KUKA KRL program: MAIN_1.src, MAIN_1.dat

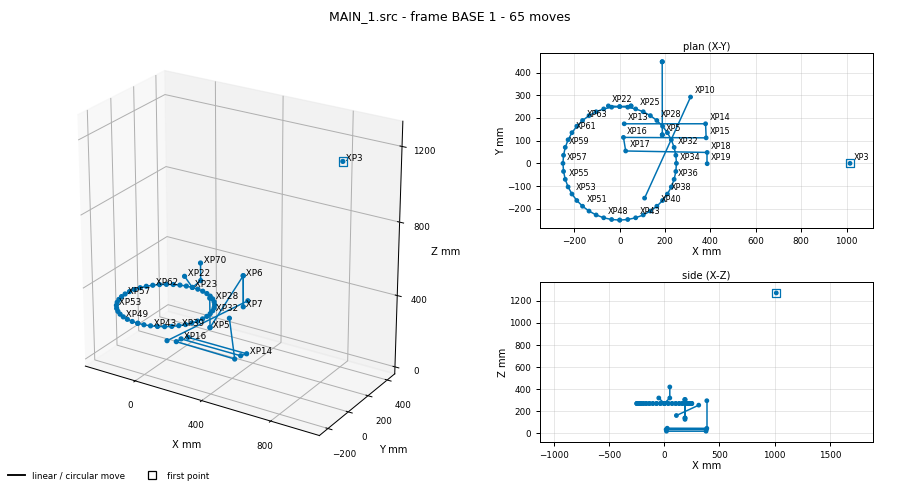
[picture p0: tool path of MAIN_1.src in frame BASE 1, 65 of 76 moves have a stored position in this frame; points joined in program order, loops and branches not executed]
--- MAIN_1.src ---
&ACCESS RVP
&REL 1
&COMMENT Generated by RoboDK
&PARAM TEMPLATE = C:\KRC\Roboter\Template\vorgabe
&PARAM EDITMASK = *
DEF MAIN_1 ( )
;FOLD INI
BAS (#INITMOV,0 )
;ENDFOLD (INI)

;FOLD STARTPOS
$BWDSTART = FALSE
PDAT_ACT = {VEL 50,ACC 100,APO_DIST 10}
BAS(#PTP_DAT)
FDAT_ACT = {TOOL_NO 0,BASE_NO 0,IPO_FRAME #BASE}
BAS (#FRAMES)
BAS (#VEL_PTP,50)
;ENDFOLD


;FOLD SET DEFAULT SPEED
$VEL.CP=0.2
BAS(#VEL_PTP,50)
BAS(#TOOL,0)
BAS(#BASE,0)
;ENDFOLD

;FOLD PTP FIRST POSITION
$BWDSTART = FALSE
PDAT_ACT = {VEL 50,ACC 100,APO_DIST 10}
FDAT_ACT = {TOOL_NO 0,BASE_NO 0,IPO_FRAME #BASE}
BAS(#FRAMES)
$ADVANCE = 5
;ENDFOLD

PTP $AXIS_ACT ; skip BCO quickly

; Program generated by RoboDK v5.6.9 for RoboDK Industrial on 26/02/2024 09:58:20
; Using nominal kinematics.
;FOLD PTP P1 Vel=100.000 % PDAT1 Tool[1] Base[1];%{PE}%R 8.3.42,%MKUKATPBASIS,%CMOVE,%VPTP,%P 1:PTP, 2:P1, 3:, 5:100, 7:PDAT1
$BWDSTART=FALSE
PDAT_ACT=PPDAT1
FDAT_ACT=FP1
BAS(#PTP_PARAMS,100)
PTP XP1 C_PTP
;ENDFOLD
;FOLD PTP P2 Vel=100.000 % PDAT2 Tool[1] Base[1];%{PE}%R 8.3.42,%MKUKATPBASIS,%CMOVE,%VPTP,%P 1:PTP, 2:P2, 3:, 5:100, 7:PDAT2
$BWDSTART=FALSE
PDAT_ACT=PPDAT2
FDAT_ACT=FP2
BAS(#PTP_PARAMS,100)
PTP XP2 C_PTP
;ENDFOLD
;FOLD LIN P3 Vel=1.000 m/s CPDAT3 Tool[1] Base[1];%{PE}%R 8.3.42,%MKUKATPBASIS,%CMOVE,%VLIN,%P 1:LIN, 2:P3, 3:, 5:1, 7:CPDAT3
$BWDSTART=FALSE
LDAT_ACT=LCPDAT3
FDAT_ACT=FP3
BAS(#CP_PARAMS,1.000)
LIN XP3 C_DIS
;ENDFOLD
$OUT[5]=TRUE
$OUT[5]=TRUE
$OUT[5]=0.5
$OUT[5]=true
$ANOUT[5]=TRUE
$ANOUT[5]=TRUE
$ANOUT[5]=0.5
$ANOUT[5]=true
var=val
var=val
WAIT FOR ($IN[5]==TRUE)
WAIT FOR ($IN[5]==TRUE)
WAIT FOR ($IN[5]==0.5)
WAIT FOR ($IN[5]==true)
START_TIMER:
$TIMER_STOP[1]=TRUE
$TIMER_FLAG[1]=FALSE
$TIMER[1]=0.100
$TIMER_STOP[1]=FALSE
WAIT FOR ($IN[5]==TRUE OR $TIMER_FLAG[1])
$TIMER_STOP[1]=TRUE
IF $TIMER_FLAG[1]== TRUE THEN
    HALT ; Timed out!
    GOTO START_TIMER
ENDIF
WAIT FOR (var==val)
START_TIMER:
$TIMER_STOP[1]=TRUE
$TIMER_FLAG[1]=FALSE
$TIMER[1]=0.100
$TIMER_STOP[1]=FALSE
WAIT FOR (var==val OR $TIMER_FLAG[1])
$TIMER_STOP[1]=TRUE
IF $TIMER_FLAG[1]== TRUE THEN
    HALT ; Timed out!
    GOTO START_TIMER
ENDIF
Wait for StrClear($LOOP_MSG[])
$LOOP_CONT = TRUE
$LOOP_MSG[] = "Message"
REMOTE_PROG_CALL_171()
CODE_INSERT_172
; Insert Comment
; ---- Setting reference (Base) ----
$BASE = {FRAME: X 719.013,Y -664.003,Z 0.000,A 0.000,B 0.000,C 0.000}
; --------------------------
; ---- Setting tool (TCP) ----
; TOOL_DATA[1] = {FRAME: X 129.073,Y 0.000,Z 85.477,A 0.000,B 22.849,C 0.000}
$TOOL = {FRAME: X 129.073,Y 0.000,Z 85.477,A 0.000,B 22.849,C 0.000}
; $TOOL = TOOL_DATA[1]
; --------------------------
$ACC.ORI1 = 800.00000
$ACC.ORI2 = 800.00000
$VEL.ORI1 = 500.00000
$VEL.ORI2 = 500.00000
$APO.CPTP = 10
$APO.CDIS = 10.000
;FOLD PTP P4 CONT Vel=100.000 % PDAT4 Tool[1] Base[1];%{PE}%R 8.3.42,%MKUKATPBASIS,%CMOVE,%VPTP,%P 1:PTP, 2:P4, 3:C_PTP, 5:100, 7:PDAT4
$BWDSTART=FALSE
PDAT_ACT=PPDAT4
FDAT_ACT=FP4
BAS(#PTP_PARAMS,100)
PTP XP4 C_PTP
;ENDFOLD
$ACC.CP = 0.20000
$VEL.CP = 0.10000
;FOLD LIN P5 Vel=0.100 m/s CPDAT5 Tool[1] Base[1];%{PE}%R 8.3.42,%MKUKATPBASIS,%CMOVE,%VLIN,%P 1:LIN, 2:P5, 3:, 5:0, 7:CPDAT5
$BWDSTART=FALSE
LDAT_ACT=LCPDAT5
FDAT_ACT=FP5
BAS(#CP_PARAMS,0.100)
LIN XP5 C_DIS
;ENDFOLD
$OUT[5]=TRUE
PICK_PART_111()
$APO.CPTP = 10
$APO.CDIS = 10.000
$ACC.CP = 0.60000
$VEL.CP = 0.30000
; Linear movement using joint targets is not supported. Change the target type to cartesian or use a joint movement.
;FOLD LIN P6 CONT Vel=0.300 m/s CPDAT6 Tool[1] Base[1];%{PE}%R 8.3.42,%MKUKATPBASIS,%CMOVE,%VLIN,%P 1:LIN, 2:P6, 3:C_DIS, 5:0, 7:CPDAT6
$BWDSTART=FALSE
LDAT_ACT=LCPDAT6
FDAT_ACT=FP6
BAS(#CP_PARAMS,0.300)
LIN XP6 C_DIS
;ENDFOLD
$ACC.CP = 0.20000
$VEL.CP = 0.10000
; MoveSearch command not implemented
;FOLD LIN P7 Vel=0.100 m/s CPDAT7 Tool[1] Base[1];%{PE}%R 8.3.42,%MKUKATPBASIS,%CMOVE,%VLIN,%P 1:LIN, 2:P7, 3:, 5:0, 7:CPDAT7
$BWDSTART=FALSE
LDAT_ACT=LCPDAT7
FDAT_ACT=FP7
BAS(#CP_PARAMS,0.100)
LIN XP7 C_DIS
;ENDFOLD
$OUT[5]=FALSE
PLACE_PART_112()
$APO.CPTP = 10
$APO.CDIS = 10.000
;FOLD LIN P8 CONT Vel=0.100 m/s CPDAT8 Tool[1] Base[1];%{PE}%R 8.3.42,%MKUKATPBASIS,%CMOVE,%VLIN,%P 1:LIN, 2:P8, 3:C_DIS, 5:0, 7:CPDAT8
$BWDSTART=FALSE
LDAT_ACT=LCPDAT8
FDAT_ACT=FP8
BAS(#CP_PARAMS,0.100)
LIN XP8 C_DIS
;ENDFOLD
; ---- Setting reference (Base) ----
$BASE = {FRAME: X 577.670,Y 392.250,Z 0.000,A 38.960,B 0.000,C 0.000}
; --------------------------
$APO.CPTP = 25
$APO.CDIS = 25.000
$ACC.ORI1 = 800.00000
$ACC.ORI2 = 800.00000
$VEL.ORI1 = 500.00000
$VEL.ORI2 = 500.00000
$ACC.CP = 0.20000
$VEL.CP = 0.10000
;FOLD PTP P9 CONT Vel=100.000 % PDAT9 Tool[1] Base[1];%{PE}%R 8.3.42,%MKUKATPBASIS,%CMOVE,%VPTP,%P 1:PTP, 2:P9, 3:C_PTP, 5:100, 7:PDAT9
$BWDSTART=FALSE
PDAT_ACT=PPDAT9
FDAT_ACT=FP9
BAS(#PTP_PARAMS,100)
PTP XP9 C_PTP
;ENDFOLD
CIRC {X 430.047,Y 43.774,Z 231.503,A -134.549,B 11.181,C 178.913},{X 109.688,Y -153.222,Z 161.073,A -134.549,B 11.181,C 178.913} C_DIS
; Circular movement using joint targets is not supported. Change the target type to cartesian or use a joint movement.
$ACC.CP = 0.20000
$VEL.CP = 0.10000
;FOLD LIN P10 Vel=0.100 m/s CPDAT10 Tool[1] Base[1];%{PE}%R 8.3.42,%MKUKATPBASIS,%CMOVE,%VLIN,%P 1:LIN, 2:P10, 3:, 5:0, 7:CPDAT10
$BWDSTART=FALSE
LDAT_ACT=LCPDAT10
FDAT_ACT=FP10
BAS(#CP_PARAMS,0.100)
LIN XP10 C_DIS
;ENDFOLD
;FOLD PTP P11 Vel=100.000 % PDAT11 Tool[1] Base[1];%{PE}%R 8.3.42,%MKUKATPBASIS,%CMOVE,%VPTP,%P 1:PTP, 2:P11, 3:, 5:100, 7:PDAT11
$BWDSTART=FALSE
PDAT_ACT=PPDAT11
FDAT_ACT=FP11
BAS(#PTP_PARAMS,100)
PTP XP11 C_PTP
;ENDFOLD
; ---- Setting reference (Base) ----
$BASE = {FRAME: X 0.000,Y 782.714,Z 377.610,A 0.000,B 0.000,C 0.000}
; --------------------------
;FOLD PTP P12 Vel=100.000 % PDAT12 Tool[1] Base[1];%{PE}%R 8.3.42,%MKUKATPBASIS,%CMOVE,%VPTP,%P 1:PTP, 2:P12, 3:, 5:100, 7:PDAT12
$BWDSTART=FALSE
PDAT_ACT=PPDAT12
FDAT_ACT=FP12
BAS(#PTP_PARAMS,100)
PTP XP12 C_PTP
;ENDFOLD
;FOLD LIN P13 Vel=0.100 m/s CPDAT13 Tool[1] Base[1];%{PE}%R 8.3.42,%MKUKATPBASIS,%CMOVE,%VLIN,%P 1:LIN, 2:P13, 3:, 5:0, 7:CPDAT13
$BWDSTART=FALSE
LDAT_ACT=LCPDAT13
FDAT_ACT=FP13
BAS(#CP_PARAMS,0.100)
LIN XP13 C_DIS
;ENDFOLD
;FOLD LIN P14 Vel=0.100 m/s CPDAT14 Tool[1] Base[1];%{PE}%R 8.3.42,%MKUKATPBASIS,%CMOVE,%VLIN,%P 1:LIN, 2:P14, 3:, 5:0, 7:CPDAT14
$BWDSTART=FALSE
LDAT_ACT=LCPDAT14
FDAT_ACT=FP14
BAS(#CP_PARAMS,0.100)
LIN XP14 C_DIS
;ENDFOLD
;FOLD LIN P15 Vel=0.100 m/s CPDAT15 Tool[1] Base[1];%{PE}%R 8.3.42,%MKUKATPBASIS,%CMOVE,%VLIN,%P 1:LIN, 2:P15, 3:, 5:0, 7:CPDAT15
$BWDSTART=FALSE
LDAT_ACT=LCPDAT15
FDAT_ACT=FP15
BAS(#CP_PARAMS,0.100)
LIN XP15 C_DIS
;ENDFOLD
;FOLD LIN P16 Vel=0.100 m/s CPDAT16 Tool[1] Base[1];%{PE}%R 8.3.42,%MKUKATPBASIS,%CMOVE,%VLIN,%P 1:LIN, 2:P16, 3:, 5:0, 7:CPDAT16
$BWDSTART=FALSE
LDAT_ACT=LCPDAT16
FDAT_ACT=FP16
BAS(#CP_PARAMS,0.100)
LIN XP16 C_DIS
;ENDFOLD
;FOLD LIN P17 Vel=0.100 m/s CPDAT17 Tool[1] Base[1];%{PE}%R 8.3.42,%MKUKATPBASIS,%CMOVE,%VLIN,%P 1:LIN, 2:P17, 3:, 5:0, 7:CPDAT17
$BWDSTART=FALSE
LDAT_ACT=LCPDAT17
FDAT_ACT=FP17
BAS(#CP_PARAMS,0.100)
LIN XP17 C_DIS
;ENDFOLD
;FOLD LIN P18 Vel=0.100 m/s CPDAT18 Tool[1] Base[1];%{PE}%R 8.3.42,%MKUKATPBASIS,%CMOVE,%VLIN,%P 1:LIN, 2:P18, 3:, 5:0, 7:CPDAT18
$BWDSTART=FALSE
LDAT_ACT=LCPDAT18
FDAT_ACT=FP18
BAS(#CP_PARAMS,0.100)
LIN XP18 C_DIS
;ENDFOLD
;FOLD LIN P19 Vel=0.100 m/s CPDAT19 Tool[1] Base[1];%{PE}%R 8.3.42,%MKUKATPBASIS,%CMOVE,%VLIN,%P 1:LIN, 2:P19, 3:, 5:0, 7:CPDAT19
$BWDSTART=FALSE
LDAT_ACT=LCPDAT19
FDAT_ACT=FP19
BAS(#CP_PARAMS,0.100)
LIN XP19 C_DIS
;ENDFOLD
;FOLD PTP P20 Vel=100.000 % PDAT20 Tool[1] Base[1];%{PE}%R 8.3.42,%MKUKATPBASIS,%CMOVE,%VPTP,%P 1:PTP, 2:P20, 3:, 5:100, 7:PDAT20
$BWDSTART=FALSE
PDAT_ACT=PPDAT20
FDAT_ACT=FP20
BAS(#PTP_PARAMS,100)
PTP XP20 C_PTP
;ENDFOLD
EVENT_PROG_START_101()
$APO.CPTP = 1
$APO.CDIS = 1.000
$VEL.CP = 1.00000
; ---- Setting reference (Base) ----
$BASE = {FRAME: X 13.637,Y -840.080,Z 0.000,A -90.000,B 0.000,C 0.000}
; --------------------------
; Show Tool 1
;FOLD PTP P21 CONT Vel=100.000 % PDAT21 Tool[1] Base[1];%{PE}%R 8.3.42,%MKUKATPBASIS,%CMOVE,%VPTP,%P 1:PTP, 2:P21, 3:C_PTP, 5:100, 7:PDAT21
$BWDSTART=FALSE
PDAT_ACT=PPDAT21
FDAT_ACT=FP21
BAS(#PTP_PARAMS,100)
PTP XP21 C_PTP
;ENDFOLD
EVENT_PATH_APPROACH_102()
;FOLD LIN P22 CONT Vel=1.000 m/s CPDAT22 Tool[1] Base[1];%{PE}%R 8.3.42,%MKUKATPBASIS,%CMOVE,%VLIN,%P 1:LIN, 2:P22, 3:C_DIS, 5:1, 7:CPDAT22
$BWDSTART=FALSE
LDAT_ACT=LCPDAT22
FDAT_ACT=FP22
BAS(#CP_PARAMS,1.000)
LIN XP22 C_DIS
;ENDFOLD
;FOLD LIN P23 CONT Vel=1.000 m/s CPDAT23 Tool[1] Base[1];%{PE}%R 8.3.42,%MKUKATPBASIS,%CMOVE,%VLIN,%P 1:LIN, 2:P23, 3:C_DIS, 5:1, 7:CPDAT23
$BWDSTART=FALSE
LDAT_ACT=LCPDAT23
FDAT_ACT=FP23
BAS(#CP_PARAMS,1.000)
LIN XP23 C_DIS
;ENDFOLD
EVENT_PATH_START_103()
$VEL.CP = 0.05000
;FOLD LIN P24 CONT Vel=0.050 m/s CPDAT24 Tool[1] Base[1];%{PE}%R 8.3.42,%MKUKATPBASIS,%CMOVE,%VLIN,%P 1:LIN, 2:P24, 3:C_DIS, 5:0, 7:CPDAT24
$BWDSTART=FALSE
LDAT_ACT=LCPDAT24
FDAT_ACT=FP24
BAS(#CP_PARAMS,0.050)
LIN XP24 C_DIS
;ENDFOLD
;FOLD LIN P25 CONT Vel=0.050 m/s CPDAT25 Tool[1] Base[1];%{PE}%R 8.3.42,%MKUKATPBASIS,%CMOVE,%VLIN,%P 1:LIN, 2:P25, 3:C_DIS, 5:0, 7:CPDAT25
$BWDSTART=FALSE
LDAT_ACT=LCPDAT25
FDAT_ACT=FP25
BAS(#CP_PARAMS,0.050)
LIN XP25 C_DIS
;ENDFOLD
;FOLD LIN P26 CONT Vel=0.050 m/s CPDAT26 Tool[1] Base[1];%{PE}%R 8.3.42,%MKUKATPBASIS,%CMOVE,%VLIN,%P 1:LIN, 2:P26, 3:C_DIS, 5:0, 7:CPDAT26
$BWDSTART=FALSE
LDAT_ACT=LCPDAT26
FDAT_ACT=FP26
BAS(#CP_PARAMS,0.050)
LIN XP26 C_DIS
;ENDFOLD
;FOLD LIN P27 CONT Vel=0.050 m/s CPDAT27 Tool[1] Base[1];%{PE}%R 8.3.42,%MKUKATPBASIS,%CMOVE,%VLIN,%P 1:LIN, 2:P27, 3:C_DIS, 5:0, 7:CPDAT27
$BWDSTART=FALSE
LDAT_ACT=LCPDAT27
FDAT_ACT=FP27
BAS(#CP_PARAMS,0.050)
LIN XP27 C_DIS
;ENDFOLD
;FOLD LIN P28 CONT Vel=0.050 m/s CPDAT28 Tool[1] Base[1];%{PE}%R 8.3.42,%MKUKATPBASIS,%CMOVE,%VLIN,%P 1:LIN, 2:P28, 3:C_DIS, 5:0, 7:CPDAT28
$BWDSTART=FALSE
LDAT_ACT=LCPDAT28
FDAT_ACT=FP28
BAS(#CP_PARAMS,0.050)
LIN XP28 C_DIS
;ENDFOLD
;FOLD LIN P29 CONT Vel=0.050 m/s CPDAT29 Tool[1] Base[1];%{PE}%R 8.3.42,%MKUKATPBASIS,%CMOVE,%VLIN,%P 1:LIN, 2:P29, 3:C_DIS, 5:0, 7:CPDAT29
$BWDSTART=FALSE
LDAT_ACT=LCPDAT29
FDAT_ACT=FP29
BAS(#CP_PARAMS,0.050)
LIN XP29 C_DIS
;ENDFOLD
;FOLD LIN P30 CONT Vel=0.050 m/s CPDAT30 Tool[1] Base[1];%{PE}%R 8.3.42,%MKUKATPBASIS,%CMOVE,%VLIN,%P 1:LIN, 2:P30, 3:C_DIS, 5:0, 7:CPDAT30
$BWDSTART=FALSE
LDAT_ACT=LCPDAT30
FDAT_ACT=FP30
BAS(#CP_PARAMS,0.050)
LIN XP30 C_DIS
;ENDFOLD
;FOLD LIN P31 CONT Vel=0.050 m/s CPDAT31 Tool[1] Base[1];%{PE}%R 8.3.42,%MKUKATPBASIS,%CMOVE,%VLIN,%P 1:LIN, 2:P31, 3:C_DIS, 5:0, 7:CPDAT31
$BWDSTART=FALSE
LDAT_ACT=LCPDAT31
FDAT_ACT=FP31
BAS(#CP_PARAMS,0.050)
LIN XP31 C_DIS
;ENDFOLD
;FOLD LIN P32 CONT Vel=0.050 m/s CPDAT32 Tool[1] Base[1];%{PE}%R 8.3.42,%MKUKATPBASIS,%CMOVE,%VLIN,%P 1:LIN, 2:P32, 3:C_DIS, 5:0, 7:CPDAT32
$BWDSTART=FALSE
LDAT_ACT=LCPDAT32
FDAT_ACT=FP32
BAS(#CP_PARAMS,0.050)
LIN XP32 C_DIS
;ENDFOLD
;FOLD LIN P33 CONT Vel=0.050 m/s CPDAT33 Tool[1] Base[1];%{PE}%R 8.3.42,%MKUKATPBASIS,%CMOVE,%VLIN,%P 1:LIN, 2:P33, 3:C_DIS, 5:0, 7:CPDAT33
$BWDSTART=FALSE
LDAT_ACT=LCPDAT33
FDAT_ACT=FP33
BAS(#CP_PARAMS,0.050)
LIN XP33 C_DIS
;ENDFOLD
;FOLD LIN P34 CONT Vel=0.050 m/s CPDAT34 Tool[1] Base[1];%{PE}%R 8.3.42,%MKUKATPBASIS,%CMOVE,%VLIN,%P 1:LIN, 2:P34, 3:C_DIS, 5:0, 7:CPDAT34
$BWDSTART=FALSE
LDAT_ACT=LCPDAT34
FDAT_ACT=FP34
BAS(#CP_PARAMS,0.050)
LIN XP34 C_DIS
;ENDFOLD
;FOLD LIN P35 CONT Vel=0.050 m/s CPDAT35 Tool[1] Base[1];%{PE}%R 8.3.42,%MKUKATPBASIS,%CMOVE,%VLIN,%P 1:LIN, 2:P35, 3:C_DIS, 5:0, 7:CPDAT35
$BWDSTART=FALSE
LDAT_ACT=LCPDAT35
FDAT_ACT=FP35
BAS(#CP_PARAMS,0.050)
LIN XP35 C_DIS
;ENDFOLD
;FOLD LIN P36 CONT Vel=0.050 m/s CPDAT36 Tool[1] Base[1];%{PE}%R 8.3.42,%MKUKATPBASIS,%CMOVE,%VLIN,%P 1:LIN, 2:P36, 3:C_DIS, 5:0, 7:CPDAT36
$BWDSTART=FALSE
LDAT_ACT=LCPDAT36
FDAT_ACT=FP36
BAS(#CP_PARAMS,0.050)
LIN XP36 C_DIS
;ENDFOLD
;FOLD LIN P37 CONT Vel=0.050 m/s CPDAT37 Tool[1] Base[1];%{PE}%R 8.3.42,%MKUKATPBASIS,%CMOVE,%VLIN,%P 1:LIN, 2:P37, 3:C_DIS, 5:0, 7:CPDAT37
$BWDSTART=FALSE
LDAT_ACT=LCPDAT37
FDAT_ACT=FP37
BAS(#CP_PARAMS,0.050)
LIN XP37 C_DIS
;ENDFOLD
;FOLD LIN P38 CONT Vel=0.050 m/s CPDAT38 Tool[1] Base[1];%{PE}%R 8.3.42,%MKUKATPBASIS,%CMOVE,%VLIN,%P 1:LIN, 2:P38, 3:C_DIS, 5:0, 7:CPDAT38
$BWDSTART=FALSE
LDAT_ACT=LCPDAT38
FDAT_ACT=FP38
BAS(#CP_PARAMS,0.050)
LIN XP38 C_DIS
;ENDFOLD
;FOLD LIN P39 CONT Vel=0.050 m/s CPDAT39 Tool[1] Base[1];%{PE}%R 8.3.42,%MKUKATPBASIS,%CMOVE,%VLIN,%P 1:LIN, 2:P39, 3:C_DIS, 5:0, 7:CPDAT39
$BWDSTART=FALSE
LDAT_ACT=LCPDAT39
FDAT_ACT=FP39
BAS(#CP_PARAMS,0.050)
LIN XP39 C_DIS
;ENDFOLD
;FOLD LIN P40 CONT Vel=0.050 m/s CPDAT40 Tool[1] Base[1];%{PE}%R 8.3.42,%MKUKATPBASIS,%CMOVE,%VLIN,%P 1:LIN, 2:P40, 3:C_DIS, 5:0, 7:CPDAT40
$BWDSTART=FALSE
LDAT_ACT=LCPDAT40
FDAT_ACT=FP40
BAS(#CP_PARAMS,0.050)
LIN XP40 C_DIS
;ENDFOLD
;FOLD LIN P41 CONT Vel=0.050 m/s CPDAT41 Tool[1] Base[1];%{PE}%R 8.3.42,%MKUKATPBASIS,%CMOVE,%VLIN,%P 1:LIN, 2:P41, 3:C_DIS, 5:0, 7:CPDAT41
$BWDSTART=FALSE
LDAT_ACT=LCPDAT41
FDAT_ACT=FP41
BAS(#CP_PARAMS,0.050)
LIN XP41 C_DIS
;ENDFOLD
;FOLD LIN P42 CONT Vel=0.050 m/s CPDAT42 Tool[1] Base[1];%{PE}%R 8.3.42,%MKUKATPBASIS,%CMOVE,%VLIN,%P 1:LIN, 2:P42, 3:C_DIS, 5:0, 7:CPDAT42
$BWDSTART=FALSE
LDAT_ACT=LCPDAT42
FDAT_ACT=FP42
BAS(#CP_PARAMS,0.050)
LIN XP42 C_DIS
;ENDFOLD
;FOLD LIN P43 CONT Vel=0.050 m/s CPDAT43 Tool[1] Base[1];%{PE}%R 8.3.42,%MKUKATPBASIS,%CMOVE,%VLIN,%P 1:LIN, 2:P43, 3:C_DIS, 5:0, 7:CPDAT43
$BWDSTART=FALSE
LDAT_ACT=LCPDAT43
FDAT_ACT=FP43
BAS(#CP_PARAMS,0.050)
LIN XP43 C_DIS
;ENDFOLD
;FOLD LIN P44 CONT Vel=0.050 m/s CPDAT44 Tool[1] Base[1];%{PE}%R 8.3.42,%MKUKATPBASIS,%CMOVE,%VLIN,%P 1:LIN, 2:P44, 3:C_DIS, 5:0, 7:CPDAT44
$BWDSTART=FALSE
LDAT_ACT=LCPDAT44
FDAT_ACT=FP44
BAS(#CP_PARAMS,0.050)
LIN XP44 C_DIS
;ENDFOLD
;FOLD LIN P45 CONT Vel=0.050 m/s CPDAT45 Tool[1] Base[1];%{PE}%R 8.3.42,%MKUKATPBASIS,%CMOVE,%VLIN,%P 1:LIN, 2:P45, 3:C_DIS, 5:0, 7:CPDAT45
$BWDSTART=FALSE
LDAT_ACT=LCPDAT45
FDAT_ACT=FP45
BAS(#CP_PARAMS,0.050)
LIN XP45 C_DIS
;ENDFOLD
;FOLD LIN P46 CONT Vel=0.050 m/s CPDAT46 Tool[1] Base[1];%{PE}%R 8.3.42,%MKUKATPBASIS,%CMOVE,%VLIN,%P 1:LIN, 2:P46, 3:C_DIS, 5:0, 7:CPDAT46
$BWDSTART=FALSE
LDAT_ACT=LCPDAT46
FDAT_ACT=FP46
BAS(#CP_PARAMS,0.050)
LIN XP46 C_DIS
;ENDFOLD
;FOLD LIN P47 CONT Vel=0.050 m/s CPDAT47 Tool[1] Base[1];%{PE}%R 8.3.42,%MKUKATPBASIS,%CMOVE,%VLIN,%P 1:LIN, 2:P47, 3:C_DIS, 5:0, 7:CPDAT47
$BWDSTART=FALSE
LDAT_ACT=LCPDAT47
FDAT_ACT=FP47
BAS(#CP_PARAMS,0.050)
LIN XP47 C_DIS
;ENDFOLD
;FOLD LIN P48 CONT Vel=0.050 m/s CPDAT48 Tool[1] Base[1];%{PE}%R 8.3.42,%MKUKATPBASIS,%CMOVE,%VLIN,%P 1:LIN, 2:P48, 3:C_DIS, 5:0, 7:CPDAT48
$BWDSTART=FALSE
LDAT_ACT=LCPDAT48
FDAT_ACT=FP48
BAS(#CP_PARAMS,0.050)
LIN XP48 C_DIS
;ENDFOLD
;FOLD LIN P49 CONT Vel=0.050 m/s CPDAT49 Tool[1] Base[1];%{PE}%R 8.3.42,%MKUKATPBASIS,%CMOVE,%VLIN,%P 1:LIN, 2:P49, 3:C_DIS, 5:0, 7:CPDAT49
$BWDSTART=FALSE
LDAT_ACT=LCPDAT49
FDAT_ACT=FP49
BAS(#CP_PARAMS,0.050)
LIN XP49 C_DIS
;ENDFOLD
;FOLD LIN P50 CONT Vel=0.050 m/s CPDAT50 Tool[1] Base[1];%{PE}%R 8.3.42,%MKUKATPBASIS,%CMOVE,%VLIN,%P 1:LIN, 2:P50, 3:C_DIS, 5:0, 7:CPDAT50
$BWDSTART=FALSE
LDAT_ACT=LCPDAT50
FDAT_ACT=FP50
BAS(#CP_PARAMS,0.050)
LIN XP50 C_DIS
;ENDFOLD
;FOLD LIN P51 CONT Vel=0.050 m/s CPDAT51 Tool[1] Base[1];%{PE}%R 8.3.42,%MKUKATPBASIS,%CMOVE,%VLIN,%P 1:LIN, 2:P51, 3:C_DIS, 5:0, 7:CPDAT51
$BWDSTART=FALSE
LDAT_ACT=LCPDAT51
FDAT_ACT=FP51
BAS(#CP_PARAMS,0.050)
LIN XP51 C_DIS
;ENDFOLD
;FOLD LIN P52 CONT Vel=0.050 m/s CPDAT52 Tool[1] Base[1];%{PE}%R 8.3.42,%MKUKATPBASIS,%CMOVE,%VLIN,%P 1:LIN, 2:P52, 3:C_DIS, 5:0, 7:CPDAT52
$BWDSTART=FALSE
LDAT_ACT=LCPDAT52
FDAT_ACT=FP52
BAS(#CP_PARAMS,0.050)
LIN XP52 C_DIS
;ENDFOLD
;FOLD LIN P53 CONT Vel=0.050 m/s CPDAT53 Tool[1] Base[1];%{PE}%R 8.3.42,%MKUKATPBASIS,%CMOVE,%VLIN,%P 1:LIN, 2:P53, 3:C_DIS, 5:0, 7:CPDAT53
$BWDSTART=FALSE
LDAT_ACT=LCPDAT53
FDAT_ACT=FP53
BAS(#CP_PARAMS,0.050)
LIN XP53 C_DIS
;ENDFOLD
;FOLD LIN P54 CONT Vel=0.050 m/s CPDAT54 Tool[1] Base[1];%{PE}%R 8.3.42,%MKUKATPBASIS,%CMOVE,%VLIN,%P 1:LIN, 2:P54, 3:C_DIS, 5:0, 7:CPDAT54
$BWDSTART=FALSE
LDAT_ACT=LCPDAT54
FDAT_ACT=FP54
BAS(#CP_PARAMS,0.050)
LIN XP54 C_DIS
;ENDFOLD
;FOLD LIN P55 CONT Vel=0.050 m/s CPDAT55 Tool[1] Base[1];%{PE}%R 8.3.42,%MKUKATPBASIS,%CMOVE,%VLIN,%P 1:LIN, 2:P55, 3:C_DIS, 5:0, 7:CPDAT55
$BWDSTART=FALSE
LDAT_ACT=LCPDAT55
FDAT_ACT=FP55
BAS(#CP_PARAMS,0.050)
LIN XP55 C_DIS
;ENDFOLD
;FOLD LIN P56 CONT Vel=0.050 m/s CPDAT56 Tool[1] Base[1];%{PE}%R 8.3.42,%MKUKATPBASIS,%CMOVE,%VLIN,%P 1:LIN, 2:P56, 3:C_DIS, 5:0, 7:CPDAT56
$BWDSTART=FALSE
LDAT_ACT=LCPDAT56
FDAT_ACT=FP56
BAS(#CP_PARAMS,0.050)
LIN XP56 C_DIS
;ENDFOLD
;FOLD LIN P57 CONT Vel=0.050 m/s CPDAT57 Tool[1] Base[1];%{PE}%R 8.3.42,%MKUKATPBASIS,%CMOVE,%VLIN,%P 1:LIN, 2:P57, 3:C_DIS, 5:0, 7:CPDAT57
$BWDSTART=FALSE
LDAT_ACT=LCPDAT57
FDAT_ACT=FP57
BAS(#CP_PARAMS,0.050)
LIN XP57 C_DIS
;ENDFOLD
;FOLD LIN P58 CONT Vel=0.050 m/s CPDAT58 Tool[1] Base[1];%{PE}%R 8.3.42,%MKUKATPBASIS,%CMOVE,%VLIN,%P 1:LIN, 2:P58, 3:C_DIS, 5:0, 7:CPDAT58
$BWDSTART=FALSE
LDAT_ACT=LCPDAT58
FDAT_ACT=FP58
BAS(#CP_PARAMS,0.050)
LIN XP58 C_DIS
;ENDFOLD
;FOLD LIN P59 CONT Vel=0.050 m/s CPDAT59 Tool[1] Base[1];%{PE}%R 8.3.42,%MKUKATPBASIS,%CMOVE,%VLIN,%P 1:LIN, 2:P59, 3:C_DIS, 5:0, 7:CPDAT59
$BWDSTART=FALSE
LDAT_ACT=LCPDAT59
FDAT_ACT=FP59
BAS(#CP_PARAMS,0.050)
LIN XP59 C_DIS
;ENDFOLD
;FOLD LIN P60 CONT Vel=0.050 m/s CPDAT60 Tool[1] Base[1];%{PE}%R 8.3.42,%MKUKATPBASIS,%CMOVE,%VLIN,%P 1:LIN, 2:P60, 3:C_DIS, 5:0, 7:CPDAT60
$BWDSTART=FALSE
LDAT_ACT=LCPDAT60
FDAT_ACT=FP60
BAS(#CP_PARAMS,0.050)
LIN XP60 C_DIS
;ENDFOLD
;FOLD LIN P61 CONT Vel=0.050 m/s CPDAT61 Tool[1] Base[1];%{PE}%R 8.3.42,%MKUKATPBASIS,%CMOVE,%VLIN,%P 1:LIN, 2:P61, 3:C_DIS, 5:0, 7:CPDAT61
$BWDSTART=FALSE
LDAT_ACT=LCPDAT61
FDAT_ACT=FP61
BAS(#CP_PARAMS,0.050)
LIN XP61 C_DIS
;ENDFOLD
;FOLD LIN P62 CONT Vel=0.050 m/s CPDAT62 Tool[1] Base[1];%{PE}%R 8.3.42,%MKUKATPBASIS,%CMOVE,%VLIN,%P 1:LIN, 2:P62, 3:C_DIS, 5:0, 7:CPDAT62
$BWDSTART=FALSE
LDAT_ACT=LCPDAT62
FDAT_ACT=FP62
BAS(#CP_PARAMS,0.050)
LIN XP62 C_DIS
;ENDFOLD
;FOLD LIN P63 CONT Vel=0.050 m/s CPDAT63 Tool[1] Base[1];%{PE}%R 8.3.42,%MKUKATPBASIS,%CMOVE,%VLIN,%P 1:LIN, 2:P63, 3:C_DIS, 5:0, 7:CPDAT63
$BWDSTART=FALSE
LDAT_ACT=LCPDAT63
FDAT_ACT=FP63
BAS(#CP_PARAMS,0.050)
LIN XP63 C_DIS
;ENDFOLD
;FOLD LIN P64 CONT Vel=0.050 m/s CPDAT64 Tool[1] Base[1];%{PE}%R 8.3.42,%MKUKATPBASIS,%CMOVE,%VLIN,%P 1:LIN, 2:P64, 3:C_DIS, 5:0, 7:CPDAT64
$BWDSTART=FALSE
LDAT_ACT=LCPDAT64
FDAT_ACT=FP64
BAS(#CP_PARAMS,0.050)
LIN XP64 C_DIS
;ENDFOLD
;FOLD LIN P65 CONT Vel=0.050 m/s CPDAT65 Tool[1] Base[1];%{PE}%R 8.3.42,%MKUKATPBASIS,%CMOVE,%VLIN,%P 1:LIN, 2:P65, 3:C_DIS, 5:0, 7:CPDAT65
$BWDSTART=FALSE
LDAT_ACT=LCPDAT65
FDAT_ACT=FP65
BAS(#CP_PARAMS,0.050)
LIN XP65 C_DIS
;ENDFOLD
;FOLD LIN P66 CONT Vel=0.050 m/s CPDAT66 Tool[1] Base[1];%{PE}%R 8.3.42,%MKUKATPBASIS,%CMOVE,%VLIN,%P 1:LIN, 2:P66, 3:C_DIS, 5:0, 7:CPDAT66
$BWDSTART=FALSE
LDAT_ACT=LCPDAT66
FDAT_ACT=FP66
BAS(#CP_PARAMS,0.050)
LIN XP66 C_DIS
;ENDFOLD
;FOLD LIN P67 CONT Vel=0.050 m/s CPDAT67 Tool[1] Base[1];%{PE}%R 8.3.42,%MKUKATPBASIS,%CMOVE,%VLIN,%P 1:LIN, 2:P67, 3:C_DIS, 5:0, 7:CPDAT67
$BWDSTART=FALSE
LDAT_ACT=LCPDAT67
FDAT_ACT=FP67
BAS(#CP_PARAMS,0.050)
LIN XP67 C_DIS
;ENDFOLD
;FOLD LIN P68 CONT Vel=0.050 m/s CPDAT68 Tool[1] Base[1];%{PE}%R 8.3.42,%MKUKATPBASIS,%CMOVE,%VLIN,%P 1:LIN, 2:P68, 3:C_DIS, 5:0, 7:CPDAT68
$BWDSTART=FALSE
LDAT_ACT=LCPDAT68
FDAT_ACT=FP68
BAS(#CP_PARAMS,0.050)
LIN XP68 C_DIS
;ENDFOLD
$VEL.CP = 1.00000
EVENT_PATH_FINISH_105()
;FOLD LIN P69 CONT Vel=1.000 m/s CPDAT69 Tool[1] Base[1];%{PE}%R 8.3.42,%MKUKATPBASIS,%CMOVE,%VLIN,%P 1:LIN, 2:P69, 3:C_DIS, 5:1, 7:CPDAT69
$BWDSTART=FALSE
LDAT_ACT=LCPDAT69
FDAT_ACT=FP69
BAS(#CP_PARAMS,1.000)
LIN XP69 C_DIS
;ENDFOLD
;FOLD LIN P70 CONT Vel=1.000 m/s CPDAT70 Tool[1] Base[1];%{PE}%R 8.3.42,%MKUKATPBASIS,%CMOVE,%VLIN,%P 1:LIN, 2:P70, 3:C_DIS, 5:1, 7:CPDAT70
$BWDSTART=FALSE
LDAT_ACT=LCPDAT70
FDAT_ACT=FP70
BAS(#CP_PARAMS,1.000)
LIN XP70 C_DIS
;ENDFOLD
EVENT_PATH_RETRACT_106()
EVENT_PROG_FINISH_107()
; ---- Setting reference (Base) ----
$BASE = {FRAME: X 719.013,Y -664.003,Z 0.000,A 0.000,B 0.000,C 0.000}
; --------------------------
;FOLD PTP P71 CONT Vel=100.000 % PDAT71 Tool[1] Base[1];%{PE}%R 8.3.42,%MKUKATPBASIS,%CMOVE,%VPTP,%P 1:PTP, 2:P71, 3:C_PTP, 5:100, 7:PDAT71
$BWDSTART=FALSE
PDAT_ACT=PPDAT71
FDAT_ACT=FP71
BAS(#PTP_PARAMS,100)
PTP XP71 C_PTP
;ENDFOLD
WAIT SEC 1.250
;FOLD LIN P72 CONT Vel=1.000 m/s CPDAT72 Tool[1] Base[1];%{PE}%R 8.3.42,%MKUKATPBASIS,%CMOVE,%VLIN,%P 1:LIN, 2:P72, 3:C_DIS, 5:1, 7:CPDAT72
$BWDSTART=FALSE
LDAT_ACT=LCPDAT72
FDAT_ACT=FP72
BAS(#CP_PARAMS,1.000)
LIN XP72 C_DIS
;ENDFOLD
WAIT FOR ($IN[1]==TRUE)
;FOLD LIN P73 CONT Vel=1.000 m/s CPDAT73 Tool[1] Base[1];%{PE}%R 8.3.42,%MKUKATPBASIS,%CMOVE,%VLIN,%P 1:LIN, 2:P73, 3:C_DIS, 5:1, 7:CPDAT73
$BWDSTART=FALSE
LDAT_ACT=LCPDAT73
FDAT_ACT=FP73
BAS(#CP_PARAMS,1.000)
LIN XP73 C_DIS
;ENDFOLD
PROG1_withaverylongnameandspecialcharacters()
END
DEF PROG1_withaverylongnameandspecialcharacters ( )
; This is a subprogram call to PROG_1
; ---- Setting reference (Base) ----
; BASE_DATA[1] = {FRAME: X 0.000,Y 1000.000,Z 0.000,A 0.000,B 0.000,C 0.000}
$BASE = {FRAME: X 0.000,Y 1000.000,Z 0.000,A 0.000,B 0.000,C 0.000}
; $BASE = BASE_DATA[1]
; --------------------------
; ---- Setting tool (TCP) ----
; TOOL_DATA[1] = {FRAME: X 0.000,Y 0.000,Z 200.000,A 0.000,B 0.000,C 0.000}
$TOOL = {FRAME: X 0.000,Y 0.000,Z 200.000,A 0.000,B 0.000,C 0.000}
; $TOOL = TOOL_DATA[1]
; --------------------------
;FOLD PTP P74 CONT Vel=100.000 % PDAT74 Tool[1] Base[1];%{PE}%R 8.3.42,%MKUKATPBASIS,%CMOVE,%VPTP,%P 1:PTP, 2:P74, 3:C_PTP, 5:100, 7:PDAT74
$BWDSTART=FALSE
PDAT_ACT=PPDAT74
FDAT_ACT=FP74
BAS(#PTP_PARAMS,100)
PTP XP74 C_PTP
;ENDFOLD
END

--- MAIN_1.dat ---
&ACCESS RVP
&REL 1
&COMMENT Generated by RoboDK
&PARAM TEMPLATE = C:\KRC\Roboter\Template\vorgabe
&PARAM EDITMASK = *
DEFDAT  MAIN_1

DECL E6AXIS XP1={AXIS: A1 -0.00000,A2 0.00000,A3 0.00000,A4 0.00000,A5 0.00000,A6 -0.00000}
DECL FDAT FP1={TOOL_NO 1,BASE_NO 1,IPO_FRAME #BASE,POINT2[] " ",TQ_STATE FALSE}
DECL PDAT PPDAT1={VEL 100.000,ACC 100.000,APO_DIST 1.000,GEAR_JERK 50.0000,EXAX_IGN 0}
DECL E6AXIS XP2={AXIS: A1 0.00000,A2 3.21124,A3 -15.42370,A4 0.00000,A5 12.21250,A6 -0.00000}
DECL FDAT FP2={TOOL_NO 1,BASE_NO 1,IPO_FRAME #BASE,POINT2[] " ",TQ_STATE FALSE}
DECL PDAT PPDAT2={VEL 100.000,ACC 100.000,APO_DIST 1.000,GEAR_JERK 50.0000,EXAX_IGN 0}
DECL E6POS XP3={X 1015.000,Y 0.000,Z 1272.000,A 0.000,B 90.000,C 0.000}
DECL FDAT FP3={TOOL_NO 1,BASE_NO 1,IPO_FRAME #BASE,POINT2[] " ",TQ_STATE FALSE}
DECL LDAT LCPDAT3={VEL 1.00000,ACC 100.000,APO_DIST 1.000,APO_FAC 50.0000,AXIS_VEL 100.000,AXIS_ACC 100.000,ORI_TYP #VAR,CIRC_TYP #BASE,JERK_FAC 50.0000,GEAR_JERK 50.0000,EXAX_IGN 0}
DECL E6AXIS XP4={AXIS: A1 -29.33220,A2 46.67700,A3 -0.02452,A4 26.54560,A5 25.39570,A6 -51.63400}
DECL FDAT FP4={TOOL_NO 1,BASE_NO 1,IPO_FRAME #BASE,POINT2[] " ",TQ_STATE FALSE}
DECL PDAT PPDAT4={VEL 100.000,ACC 100.000,APO_DIST 10.000,GEAR_JERK 50.0000,EXAX_IGN 0}
DECL E6POS XP5={X 187.786,Y 125.499,Z 139.112,A -179.997,B 0.180,C 179.996}
DECL FDAT FP5={TOOL_NO 1,BASE_NO 1,IPO_FRAME #BASE,POINT2[] " ",TQ_STATE FALSE}
DECL LDAT LCPDAT5={VEL 0.10000,ACC 100.000,APO_DIST 1.000,APO_FAC 50.0000,AXIS_VEL 100.000,AXIS_ACC 100.000,ORI_TYP #VAR,CIRC_TYP #BASE,JERK_FAC 50.0000,GEAR_JERK 50.0000,EXAX_IGN 0}
DECL E6POS XP6={X 187.272,Y 447.522,Z 305.347,A 179.999,B 0.185,C -179.998}
DECL FDAT FP6={TOOL_NO 1,BASE_NO 1,IPO_FRAME #BASE,POINT2[] " ",TQ_STATE FALSE}
DECL LDAT LCPDAT6={VEL 0.30000,ACC 100.000,APO_DIST 10.000,APO_FAC 50.0000,AXIS_VEL 100.000,AXIS_ACC 100.000,ORI_TYP #VAR,CIRC_TYP #BASE,JERK_FAC 50.0000,GEAR_JERK 50.0000,EXAX_IGN 0}
DECL E6POS XP7={X 187.851,Y 447.517,Z 126.235,A 179.999,B 0.185,C -179.998}
DECL FDAT FP7={TOOL_NO 1,BASE_NO 1,IPO_FRAME #BASE,POINT2[] " ",TQ_STATE FALSE}
DECL LDAT LCPDAT7={VEL 0.10000,ACC 100.000,APO_DIST 1.000,APO_FAC 50.0000,AXIS_VEL 100.000,AXIS_ACC 100.000,ORI_TYP #VAR,CIRC_TYP #BASE,JERK_FAC 50.0000,GEAR_JERK 50.0000,EXAX_IGN 0}
DECL E6POS XP8={X 187.272,Y 447.522,Z 305.347,A 179.999,B 0.185,C -179.998}
DECL FDAT FP8={TOOL_NO 1,BASE_NO 1,IPO_FRAME #BASE,POINT2[] " ",TQ_STATE FALSE}
DECL LDAT LCPDAT8={VEL 0.10000,ACC 100.000,APO_DIST 10.000,APO_FAC 50.0000,AXIS_VEL 100.000,AXIS_ACC 100.000,ORI_TYP #VAR,CIRC_TYP #BASE,JERK_FAC 50.0000,GEAR_JERK 50.0000,EXAX_IGN 0}
DECL E6AXIS XP9={AXIS: A1 52.18600,A2 45.67580,A3 6.92000,A4 66.73420,A5 19.93230,A6 -92.73000}
DECL FDAT FP9={TOOL_NO 1,BASE_NO 1,IPO_FRAME #BASE,POINT2[] " ",TQ_STATE FALSE}
DECL PDAT PPDAT9={VEL 100.000,ACC 100.000,APO_DIST 25.000,GEAR_JERK 50.0000,EXAX_IGN 0}
DECL E6POS XP10={X 312.208,Y 292.214,Z 255.156,A -134.549,B 11.181,C 178.913}
DECL FDAT FP10={TOOL_NO 1,BASE_NO 1,IPO_FRAME #BASE,POINT2[] " ",TQ_STATE FALSE}
DECL LDAT LCPDAT10={VEL 0.10000,ACC 100.000,APO_DIST 1.000,APO_FAC 50.0000,AXIS_VEL 100.000,AXIS_ACC 100.000,ORI_TYP #VAR,CIRC_TYP #BASE,JERK_FAC 50.0000,GEAR_JERK 50.0000,EXAX_IGN 0}
DECL E6AXIS XP11={AXIS: A1 -0.00000,A2 0.00000,A3 0.00000,A4 0.00000,A5 0.00000,A6 -0.00000}
DECL FDAT FP11={TOOL_NO 1,BASE_NO 1,IPO_FRAME #BASE,POINT2[] " ",TQ_STATE FALSE}
DECL PDAT PPDAT11={VEL 100.000,ACC 100.000,APO_DIST 1.000,GEAR_JERK 50.0000,EXAX_IGN 0}
DECL E6AXIS XP12={AXIS: A1 88.67600,A2 29.60160,A3 -6.42883,A4 -1.98422,A5 49.47920,A6 4.54769}
DECL FDAT FP12={TOOL_NO 1,BASE_NO 1,IPO_FRAME #BASE,POINT2[] " ",TQ_STATE FALSE}
DECL PDAT PPDAT12={VEL 100.000,ACC 100.000,APO_DIST 1.000,GEAR_JERK 50.0000,EXAX_IGN 0}
DECL E6POS XP13={X 19.898,Y 174.307,Z 19.008,A -94.928,B -5.426,C -179.533}
DECL FDAT FP13={TOOL_NO 1,BASE_NO 1,IPO_FRAME #BASE,POINT2[] " ",TQ_STATE FALSE}
DECL LDAT LCPDAT13={VEL 0.10000,ACC 100.000,APO_DIST 1.000,APO_FAC 50.0000,AXIS_VEL 100.000,AXIS_ACC 100.000,ORI_TYP #VAR,CIRC_TYP #BASE,JERK_FAC 50.0000,GEAR_JERK 50.0000,EXAX_IGN 0}
DECL E6POS XP14={X 378.402,Y 174.416,Z 18.997,A -94.928,B -5.426,C -179.533}
DECL FDAT FP14={TOOL_NO 1,BASE_NO 1,IPO_FRAME #BASE,POINT2[] " ",TQ_STATE FALSE}
DECL LDAT LCPDAT14={VEL 0.10000,ACC 100.000,APO_DIST 1.000,APO_FAC 50.0000,AXIS_VEL 100.000,AXIS_ACC 100.000,ORI_TYP #VAR,CIRC_TYP #BASE,JERK_FAC 50.0000,GEAR_JERK 50.0000,EXAX_IGN 0}
DECL E6POS XP15={X 380.996,Y 112.363,Z 34.882,A -95.294,B -18.136,C -178.348}
DECL FDAT FP15={TOOL_NO 1,BASE_NO 1,IPO_FRAME #BASE,POINT2[] " ",TQ_STATE FALSE}
DECL LDAT LCPDAT15={VEL 0.10000,ACC 100.000,APO_DIST 1.000,APO_FAC 50.0000,AXIS_VEL 100.000,AXIS_ACC 100.000,ORI_TYP #VAR,CIRC_TYP #BASE,JERK_FAC 50.0000,GEAR_JERK 50.0000,EXAX_IGN 0}
DECL E6POS XP16={X 16.551,Y 114.359,Z 34.226,A -95.294,B -18.136,C -178.348}
DECL FDAT FP16={TOOL_NO 1,BASE_NO 1,IPO_FRAME #BASE,POINT2[] " ",TQ_STATE FALSE}
DECL LDAT LCPDAT16={VEL 0.10000,ACC 100.000,APO_DIST 1.000,APO_FAC 50.0000,AXIS_VEL 100.000,AXIS_ACC 100.000,ORI_TYP #VAR,CIRC_TYP #BASE,JERK_FAC 50.0000,GEAR_JERK 50.0000,EXAX_IGN 0}
DECL E6POS XP17={X 26.434,Y 54.524,Z 46.072,A -95.461,B 4.348,C 179.585}
DECL FDAT FP17={TOOL_NO 1,BASE_NO 1,IPO_FRAME #BASE,POINT2[] " ",TQ_STATE FALSE}
DECL LDAT LCPDAT17={VEL 0.10000,ACC 100.000,APO_DIST 1.000,APO_FAC 50.0000,AXIS_VEL 100.000,AXIS_ACC 100.000,ORI_TYP #VAR,CIRC_TYP #BASE,JERK_FAC 50.0000,GEAR_JERK 50.0000,EXAX_IGN 0}
DECL E6POS XP18={X 385.448,Y 48.050,Z 45.137,A -95.590,B 11.181,C 178.913}
DECL FDAT FP18={TOOL_NO 1,BASE_NO 1,IPO_FRAME #BASE,POINT2[] " ",TQ_STATE FALSE}
DECL LDAT LCPDAT18={VEL 0.10000,ACC 100.000,APO_DIST 1.000,APO_FAC 50.0000,AXIS_VEL 100.000,AXIS_ACC 100.000,ORI_TYP #VAR,CIRC_TYP #BASE,JERK_FAC 50.0000,GEAR_JERK 50.0000,EXAX_IGN 0}
DECL E6POS XP19={X 385.448,Y -1.625,Z 295.251,A -95.590,B 11.181,C 178.913}
DECL FDAT FP19={TOOL_NO 1,BASE_NO 1,IPO_FRAME #BASE,POINT2[] " ",TQ_STATE FALSE}
DECL LDAT LCPDAT19={VEL 0.10000,ACC 100.000,APO_DIST 1.000,APO_FAC 50.0000,AXIS_VEL 100.000,AXIS_ACC 100.000,ORI_TYP #VAR,CIRC_TYP #BASE,JERK_FAC 50.0000,GEAR_JERK 50.0000,EXAX_IGN 0}
DECL E6AXIS XP20={AXIS: A1 -0.00000,A2 0.00000,A3 0.00000,A4 0.00000,A5 0.00000,A6 -0.00000}
DECL FDAT FP20={TOOL_NO 1,BASE_NO 1,IPO_FRAME #BASE,POINT2[] " ",TQ_STATE FALSE}
DECL PDAT PPDAT20={VEL 100.000,ACC 100.000,APO_DIST 1.000,GEAR_JERK 50.0000,EXAX_IGN 0}
DECL E6AXIS XP21={AXIS: A1 -68.09030,A2 24.20190,A3 26.78550,A4 38.21340,A5 36.20170,A6 -98.79640}
DECL FDAT FP21={TOOL_NO 1,BASE_NO 1,IPO_FRAME #BASE,POINT2[] " ",TQ_STATE FALSE}
DECL PDAT PPDAT21={VEL 100.000,ACC 100.000,APO_DIST 1.000,GEAR_JERK 50.0000,EXAX_IGN 0}
DECL E6POS XP22={X -49.895,Y 253.259,Z 319.999,A -90.000,B 0.353,C -179.975}
DECL FDAT FP22={TOOL_NO 1,BASE_NO 1,IPO_FRAME #BASE,POINT2[] " ",TQ_STATE FALSE}
DECL LDAT LCPDAT22={VEL 1.00000,ACC 100.000,APO_DIST 1.000,APO_FAC 50.0000,AXIS_VEL 100.000,AXIS_ACC 100.000,ORI_TYP #VAR,CIRC_TYP #BASE,JERK_FAC 50.0000,GEAR_JERK 50.0000,EXAX_IGN 0}
DECL E6POS XP23={X 0.000,Y 250.000,Z 270.000,A -90.000,B 0.353,C -179.975}
DECL FDAT FP23={TOOL_NO 1,BASE_NO 1,IPO_FRAME #BASE,POINT2[] " ",TQ_STATE FALSE}
DECL LDAT LCPDAT23={VEL 1.00000,ACC 100.000,APO_DIST 1.000,APO_FAC 50.0000,AXIS_VEL 100.000,AXIS_ACC 100.000,ORI_TYP #VAR,CIRC_TYP #BASE,JERK_FAC 50.0000,GEAR_JERK 50.0000,EXAX_IGN 0}
DECL E6POS XP24={X 35.579,Y 247.455,Z 270.000,A -90.000,B 0.345,C -179.925}
DECL FDAT FP24={TOOL_NO 1,BASE_NO 1,IPO_FRAME #BASE,POINT2[] " ",TQ_STATE FALSE}
DECL LDAT LCPDAT24={VEL 0.05000,ACC 100.000,APO_DIST 1.000,APO_FAC 50.0000,AXIS_VEL 100.000,AXIS_ACC 100.000,ORI_TYP #VAR,CIRC_TYP #BASE,JERK_FAC 50.0000,GEAR_JERK 50.0000,EXAX_IGN 0}
DECL E6POS XP25={X 70.433,Y 239.873,Z 270.000,A -89.999,B 0.331,C -179.876}
DECL FDAT FP25={TOOL_NO 1,BASE_NO 1,IPO_FRAME #BASE,POINT2[] " ",TQ_STATE FALSE}
DECL LDAT LCPDAT25={VEL 0.05000,ACC 100.000,APO_DIST 1.000,APO_FAC 50.0000,AXIS_VEL 100.000,AXIS_ACC 100.000,ORI_TYP #VAR,CIRC_TYP #BASE,JERK_FAC 50.0000,GEAR_JERK 50.0000,EXAX_IGN 0}
DECL E6POS XP26={X 103.854,Y 227.408,Z 270.000,A -89.999,B 0.310,C -179.831}
DECL FDAT FP26={TOOL_NO 1,BASE_NO 1,IPO_FRAME #BASE,POINT2[] " ",TQ_STATE FALSE}
DECL LDAT LCPDAT26={VEL 0.05000,ACC 100.000,APO_DIST 1.000,APO_FAC 50.0000,AXIS_VEL 100.000,AXIS_ACC 100.000,ORI_TYP #VAR,CIRC_TYP #BASE,JERK_FAC 50.0000,GEAR_JERK 50.0000,EXAX_IGN 0}
DECL E6POS XP27={X 135.160,Y 210.313,Z 270.000,A -89.999,B 0.283,C -179.788}
DECL FDAT FP27={TOOL_NO 1,BASE_NO 1,IPO_FRAME #BASE,POINT2[] " ",TQ_STATE FALSE}
DECL LDAT LCPDAT27={VEL 0.05000,ACC 100.000,APO_DIST 1.000,APO_FAC 50.0000,AXIS_VEL 100.000,AXIS_ACC 100.000,ORI_TYP #VAR,CIRC_TYP #BASE,JERK_FAC 50.0000,GEAR_JERK 50.0000,EXAX_IGN 0}
DECL E6POS XP28={X 163.715,Y 188.937,Z 270.000,A -89.999,B 0.250,C -179.750}
DECL FDAT FP28={TOOL_NO 1,BASE_NO 1,IPO_FRAME #BASE,POINT2[] " ",TQ_STATE FALSE}
DECL LDAT LCPDAT28={VEL 0.05000,ACC 100.000,APO_DIST 1.000,APO_FAC 50.0000,AXIS_VEL 100.000,AXIS_ACC 100.000,ORI_TYP #VAR,CIRC_TYP #BASE,JERK_FAC 50.0000,GEAR_JERK 50.0000,EXAX_IGN 0}
DECL E6POS XP29={X 188.937,Y 163.715,Z 270.000,A -89.999,B 0.212,C -179.717}
DECL FDAT FP29={TOOL_NO 1,BASE_NO 1,IPO_FRAME #BASE,POINT2[] " ",TQ_STATE FALSE}
DECL LDAT LCPDAT29={VEL 0.05000,ACC 100.000,APO_DIST 1.000,APO_FAC 50.0000,AXIS_VEL 100.000,AXIS_ACC 100.000,ORI_TYP #VAR,CIRC_TYP #BASE,JERK_FAC 50.0000,GEAR_JERK 50.0000,EXAX_IGN 0}
DECL E6POS XP30={X 210.313,Y 135.160,Z 270.000,A -89.999,B 0.170,C -179.689}
DECL FDAT FP30={TOOL_NO 1,BASE_NO 1,IPO_FRAME #BASE,POINT2[] " ",TQ_STATE FALSE}
DECL LDAT LCPDAT30={VEL 0.05000,ACC 100.000,APO_DIST 1.000,APO_FAC 50.0000,AXIS_VEL 100.000,AXIS_ACC 100.000,ORI_TYP #VAR,CIRC_TYP #BASE,JERK_FAC 50.0000,GEAR_JERK 50.0000,EXAX_IGN 0}
DECL E6POS XP31={X 227.408,Y 103.854,Z 270.000,A -89.999,B 0.124,C -179.668}
DECL FDAT FP31={TOOL_NO 1,BASE_NO 1,IPO_FRAME #BASE,POINT2[] " ",TQ_STATE FALSE}
DECL LDAT LCPDAT31={VEL 0.05000,ACC 100.000,APO_DIST 1.000,APO_FAC 50.0000,AXIS_VEL 100.000,AXIS_ACC 100.000,ORI_TYP #VAR,CIRC_TYP #BASE,JERK_FAC 50.0000,GEAR_JERK 50.0000,EXAX_IGN 0}
DECL E6POS XP32={X 239.873,Y 70.433,Z 270.000,A -90.000,B 0.075,C -179.654}
DECL FDAT FP32={TOOL_NO 1,BASE_NO 1,IPO_FRAME #BASE,POINT2[] " ",TQ_STATE FALSE}
DECL LDAT LCPDAT32={VEL 0.05000,ACC 100.000,APO_DIST 1.000,APO_FAC 50.0000,AXIS_VEL 100.000,AXIS_ACC 100.000,ORI_TYP #VAR,CIRC_TYP #BASE,JERK_FAC 50.0000,GEAR_JERK 50.0000,EXAX_IGN 0}
DECL E6POS XP33={X 247.455,Y 35.579,Z 270.000,A -90.000,B 0.025,C -179.647}
DECL FDAT FP33={TOOL_NO 1,BASE_NO 1,IPO_FRAME #BASE,POINT2[] " ",TQ_STATE FALSE}
DECL LDAT LCPDAT33={VEL 0.05000,ACC 100.000,APO_DIST 1.000,APO_FAC 50.0000,AXIS_VEL 100.000,AXIS_ACC 100.000,ORI_TYP #VAR,CIRC_TYP #BASE,JERK_FAC 50.0000,GEAR_JERK 50.0000,EXAX_IGN 0}
DECL E6POS XP34={X 250.000,Y 0.000,Z 270.000,A -90.000,B -0.025,C -179.647}
DECL FDAT FP34={TOOL_NO 1,BASE_NO 1,IPO_FRAME #BASE,POINT2[] " ",TQ_STATE FALSE}
DECL LDAT LCPDAT34={VEL 0.05000,ACC 100.000,APO_DIST 1.000,APO_FAC 50.0000,AXIS_VEL 100.000,AXIS_ACC 100.000,ORI_TYP #VAR,CIRC_TYP #BASE,JERK_FAC 50.0000,GEAR_JERK 50.0000,EXAX_IGN 0}
DECL E6POS XP35={X 247.455,Y -35.579,Z 270.000,A -90.000,B -0.075,C -179.654}
DECL FDAT FP35={TOOL_NO 1,BASE_NO 1,IPO_FRAME #BASE,POINT2[] " ",TQ_STATE FALSE}
DECL LDAT LCPDAT35={VEL 0.05000,ACC 100.000,APO_DIST 1.000,APO_FAC 50.0000,AXIS_VEL 100.000,AXIS_ACC 100.000,ORI_TYP #VAR,CIRC_TYP #BASE,JERK_FAC 50.0000,GEAR_JERK 50.0000,EXAX_IGN 0}
DECL E6POS XP36={X 239.873,Y -70.433,Z 270.000,A -90.001,B -0.124,C -179.668}
DECL FDAT FP36={TOOL_NO 1,BASE_NO 1,IPO_FRAME #BASE,POINT2[] " ",TQ_STATE FALSE}
DECL LDAT LCPDAT36={VEL 0.05000,ACC 100.000,APO_DIST 1.000,APO_FAC 50.0000,AXIS_VEL 100.000,AXIS_ACC 100.000,ORI_TYP #VAR,CIRC_TYP #BASE,JERK_FAC 50.0000,GEAR_JERK 50.0000,EXAX_IGN 0}
DECL E6POS XP37={X 227.408,Y -103.854,Z 270.000,A -90.001,B -0.170,C -179.689}
DECL FDAT FP37={TOOL_NO 1,BASE_NO 1,IPO_FRAME #BASE,POINT2[] " ",TQ_STATE FALSE}
DECL LDAT LCPDAT37={VEL 0.05000,ACC 100.000,APO_DIST 1.000,APO_FAC 50.0000,AXIS_VEL 100.000,AXIS_ACC 100.000,ORI_TYP #VAR,CIRC_TYP #BASE,JERK_FAC 50.0000,GEAR_JERK 50.0000,EXAX_IGN 0}
DECL E6POS XP38={X 210.313,Y -135.160,Z 270.000,A -90.001,B -0.212,C -179.717}
DECL FDAT FP38={TOOL_NO 1,BASE_NO 1,IPO_FRAME #BASE,POINT2[] " ",TQ_STATE FALSE}
DECL LDAT LCPDAT38={VEL 0.05000,ACC 100.000,APO_DIST 1.000,APO_FAC 50.0000,AXIS_VEL 100.000,AXIS_ACC 100.000,ORI_TYP #VAR,CIRC_TYP #BASE,JERK_FAC 50.0000,GEAR_JERK 50.0000,EXAX_IGN 0}
DECL E6POS XP39={X 188.937,Y -163.715,Z 270.000,A -90.001,B -0.250,C -179.750}
DECL FDAT FP39={TOOL_NO 1,BASE_NO 1,IPO_FRAME #BASE,POINT2[] " ",TQ_STATE FALSE}
DECL LDAT LCPDAT39={VEL 0.05000,ACC 100.000,APO_DIST 1.000,APO_FAC 50.0000,AXIS_VEL 100.000,AXIS_ACC 100.000,ORI_TYP #VAR,CIRC_TYP #BASE,JERK_FAC 50.0000,GEAR_JERK 50.0000,EXAX_IGN 0}
DECL E6POS XP40={X 163.715,Y -188.937,Z 270.000,A -90.001,B -0.283,C -179.788}
DECL FDAT FP40={TOOL_NO 1,BASE_NO 1,IPO_FRAME #BASE,POINT2[] " ",TQ_STATE FALSE}
DECL LDAT LCPDAT40={VEL 0.05000,ACC 100.000,APO_DIST 1.000,APO_FAC 50.0000,AXIS_VEL 100.000,AXIS_ACC 100.000,ORI_TYP #VAR,CIRC_TYP #BASE,JERK_FAC 50.0000,GEAR_JERK 50.0000,EXAX_IGN 0}
DECL E6POS XP41={X 135.160,Y -210.313,Z 270.000,A -90.001,B -0.311,C -179.830}
DECL FDAT FP41={TOOL_NO 1,BASE_NO 1,IPO_FRAME #BASE,POINT2[] " ",TQ_STATE FALSE}
DECL LDAT LCPDAT41={VEL 0.05000,ACC 100.000,APO_DIST 1.000,APO_FAC 50.0000,AXIS_VEL 100.000,AXIS_ACC 100.000,ORI_TYP #VAR,CIRC_TYP #BASE,JERK_FAC 50.0000,GEAR_JERK 50.0000,EXAX_IGN 0}
DECL E6POS XP42={X 103.854,Y -227.408,Z 270.000,A -90.001,B -0.332,C -179.876}
DECL FDAT FP42={TOOL_NO 1,BASE_NO 1,IPO_FRAME #BASE,POINT2[] " ",TQ_STATE FALSE}
DECL LDAT LCPDAT42={VEL 0.05000,ACC 100.000,APO_DIST 1.000,APO_FAC 50.0000,AXIS_VEL 100.000,AXIS_ACC 100.000,ORI_TYP #VAR,CIRC_TYP #BASE,JERK_FAC 50.0000,GEAR_JERK 50.0000,EXAX_IGN 0}
DECL E6POS XP43={X 70.433,Y -239.873,Z 270.000,A -90.000,B -0.346,C -179.925}
DECL FDAT FP43={TOOL_NO 1,BASE_NO 1,IPO_FRAME #BASE,POINT2[] " ",TQ_STATE FALSE}
DECL LDAT LCPDAT43={VEL 0.05000,ACC 100.000,APO_DIST 1.000,APO_FAC 50.0000,AXIS_VEL 100.000,AXIS_ACC 100.000,ORI_TYP #VAR,CIRC_TYP #BASE,JERK_FAC 50.0000,GEAR_JERK 50.0000,EXAX_IGN 0}
DECL E6POS XP44={X 35.579,Y -247.455,Z 270.000,A -90.000,B -0.353,C -179.975}
DECL FDAT FP44={TOOL_NO 1,BASE_NO 1,IPO_FRAME #BASE,POINT2[] " ",TQ_STATE FALSE}
DECL LDAT LCPDAT44={VEL 0.05000,ACC 100.000,APO_DIST 1.000,APO_FAC 50.0000,AXIS_VEL 100.000,AXIS_ACC 100.000,ORI_TYP #VAR,CIRC_TYP #BASE,JERK_FAC 50.0000,GEAR_JERK 50.0000,EXAX_IGN 0}
DECL E6POS XP45={X 0.000,Y -250.000,Z 270.000,A -90.000,B -0.353,C -179.975}
DECL FDAT FP45={TOOL_NO 1,BASE_NO 1,IPO_FRAME #BASE,POINT2[] " ",TQ_STATE FALSE}
DECL LDAT LCPDAT45={VEL 0.05000,ACC 100.000,APO_DIST 1.000,APO_FAC 50.0000,AXIS_VEL 100.000,AXIS_ACC 100.000,ORI_TYP #VAR,CIRC_TYP #BASE,JERK_FAC 50.0000,GEAR_JERK 50.0000,EXAX_IGN 0}
DECL E6POS XP46={X 0.000,Y -250.000,Z 270.000,A -90.000,B -0.353,C 179.975}
DECL FDAT FP46={TOOL_NO 1,BASE_NO 1,IPO_FRAME #BASE,POINT2[] " ",TQ_STATE FALSE}
DECL LDAT LCPDAT46={VEL 0.05000,ACC 100.000,APO_DIST 1.000,APO_FAC 50.0000,AXIS_VEL 100.000,AXIS_ACC 100.000,ORI_TYP #VAR,CIRC_TYP #BASE,JERK_FAC 50.0000,GEAR_JERK 50.0000,EXAX_IGN 0}
DECL E6POS XP47={X -35.579,Y -247.455,Z 270.000,A -90.000,B -0.346,C 179.925}
DECL FDAT FP47={TOOL_NO 1,BASE_NO 1,IPO_FRAME #BASE,POINT2[] " ",TQ_STATE FALSE}
DECL LDAT LCPDAT47={VEL 0.05000,ACC 100.000,APO_DIST 1.000,APO_FAC 50.0000,AXIS_VEL 100.000,AXIS_ACC 100.000,ORI_TYP #VAR,CIRC_TYP #BASE,JERK_FAC 50.0000,GEAR_JERK 50.0000,EXAX_IGN 0}
DECL E6POS XP48={X -70.433,Y -239.873,Z 270.000,A -89.999,B -0.331,C 179.876}
DECL FDAT FP48={TOOL_NO 1,BASE_NO 1,IPO_FRAME #BASE,POINT2[] " ",TQ_STATE FALSE}
DECL LDAT LCPDAT48={VEL 0.05000,ACC 100.000,APO_DIST 1.000,APO_FAC 50.0000,AXIS_VEL 100.000,AXIS_ACC 100.000,ORI_TYP #VAR,CIRC_TYP #BASE,JERK_FAC 50.0000,GEAR_JERK 50.0000,EXAX_IGN 0}
DECL E6POS XP49={X -103.854,Y -227.408,Z 270.000,A -89.999,B -0.310,C 179.831}
DECL FDAT FP49={TOOL_NO 1,BASE_NO 1,IPO_FRAME #BASE,POINT2[] " ",TQ_STATE FALSE}
DECL LDAT LCPDAT49={VEL 0.05000,ACC 100.000,APO_DIST 1.000,APO_FAC 50.0000,AXIS_VEL 100.000,AXIS_ACC 100.000,ORI_TYP #VAR,CIRC_TYP #BASE,JERK_FAC 50.0000,GEAR_JERK 50.0000,EXAX_IGN 0}
DECL E6POS XP50={X -135.160,Y -210.313,Z 270.000,A -89.999,B -0.283,C 179.788}
DECL FDAT FP50={TOOL_NO 1,BASE_NO 1,IPO_FRAME #BASE,POINT2[] " ",TQ_STATE FALSE}
DECL LDAT LCPDAT50={VEL 0.05000,ACC 100.000,APO_DIST 1.000,APO_FAC 50.0000,AXIS_VEL 100.000,AXIS_ACC 100.000,ORI_TYP #VAR,CIRC_TYP #BASE,JERK_FAC 50.0000,GEAR_JERK 50.0000,EXAX_IGN 0}
DECL E6POS XP51={X -163.715,Y -188.937,Z 270.000,A -89.999,B -0.250,C 179.750}
DECL FDAT FP51={TOOL_NO 1,BASE_NO 1,IPO_FRAME #BASE,POINT2[] " ",TQ_STATE FALSE}
DECL LDAT LCPDAT51={VEL 0.05000,ACC 100.000,APO_DIST 1.000,APO_FAC 50.0000,AXIS_VEL 100.000,AXIS_ACC 100.000,ORI_TYP #VAR,CIRC_TYP #BASE,JERK_FAC 50.0000,GEAR_JERK 50.0000,EXAX_IGN 0}
DECL E6POS XP52={X -188.937,Y -163.715,Z 270.000,A -89.999,B -0.212,C 179.717}
DECL FDAT FP52={TOOL_NO 1,BASE_NO 1,IPO_FRAME #BASE,POINT2[] " ",TQ_STATE FALSE}
DECL LDAT LCPDAT52={VEL 0.05000,ACC 100.000,APO_DIST 1.000,APO_FAC 50.0000,AXIS_VEL 100.000,AXIS_ACC 100.000,ORI_TYP #VAR,CIRC_TYP #BASE,JERK_FAC 50.0000,GEAR_JERK 50.0000,EXAX_IGN 0}
DECL E6POS XP53={X -210.313,Y -135.160,Z 270.000,A -89.999,B -0.169,C 179.690}
DECL FDAT FP53={TOOL_NO 1,BASE_NO 1,IPO_FRAME #BASE,POINT2[] " ",TQ_STATE FALSE}
DECL LDAT LCPDAT53={VEL 0.05000,ACC 100.000,APO_DIST 1.000,APO_FAC 50.0000,AXIS_VEL 100.000,AXIS_ACC 100.000,ORI_TYP #VAR,CIRC_TYP #BASE,JERK_FAC 50.0000,GEAR_JERK 50.0000,EXAX_IGN 0}
DECL E6POS XP54={X -227.408,Y -103.854,Z 270.000,A -89.999,B -0.123,C 179.669}
DECL FDAT FP54={TOOL_NO 1,BASE_NO 1,IPO_FRAME #BASE,POINT2[] " ",TQ_STATE FALSE}
DECL LDAT LCPDAT54={VEL 0.05000,ACC 100.000,APO_DIST 1.000,APO_FAC 50.0000,AXIS_VEL 100.000,AXIS_ACC 100.000,ORI_TYP #VAR,CIRC_TYP #BASE,JERK_FAC 50.0000,GEAR_JERK 50.0000,EXAX_IGN 0}
DECL E6POS XP55={X -239.873,Y -70.433,Z 270.000,A -90.000,B -0.075,C 179.654}
DECL FDAT FP55={TOOL_NO 1,BASE_NO 1,IPO_FRAME #BASE,POINT2[] " ",TQ_STATE FALSE}
DECL LDAT LCPDAT55={VEL 0.05000,ACC 100.000,APO_DIST 1.000,APO_FAC 50.0000,AXIS_VEL 100.000,AXIS_ACC 100.000,ORI_TYP #VAR,CIRC_TYP #BASE,JERK_FAC 50.0000,GEAR_JERK 50.0000,EXAX_IGN 0}
DECL E6POS XP56={X -247.455,Y -35.579,Z 270.000,A -90.000,B -0.025,C 179.647}
DECL FDAT FP56={TOOL_NO 1,BASE_NO 1,IPO_FRAME #BASE,POINT2[] " ",TQ_STATE FALSE}
DECL LDAT LCPDAT56={VEL 0.05000,ACC 100.000,APO_DIST 1.000,APO_FAC 50.0000,AXIS_VEL 100.000,AXIS_ACC 100.000,ORI_TYP #VAR,CIRC_TYP #BASE,JERK_FAC 50.0000,GEAR_JERK 50.0000,EXAX_IGN 0}
DECL E6POS XP57={X -250.000,Y 0.000,Z 270.000,A -90.000,B 0.025,C 179.647}
DECL FDAT FP57={TOOL_NO 1,BASE_NO 1,IPO_FRAME #BASE,POINT2[] " ",TQ_STATE FALSE}
DECL LDAT LCPDAT57={VEL 0.05000,ACC 100.000,APO_DIST 1.000,APO_FAC 50.0000,AXIS_VEL 100.000,AXIS_ACC 100.000,ORI_TYP #VAR,CIRC_TYP #BASE,JERK_FAC 50.0000,GEAR_JERK 50.0000,EXAX_IGN 0}
DECL E6POS XP58={X -247.455,Y 35.579,Z 270.000,A -90.000,B 0.075,C 179.655}
DECL FDAT FP58={TOOL_NO 1,BASE_NO 1,IPO_FRAME #BASE,POINT2[] " ",TQ_STATE FALSE}
DECL LDAT LCPDAT58={VEL 0.05000,ACC 100.000,APO_DIST 1.000,APO_FAC 50.0000,AXIS_VEL 100.000,AXIS_ACC 100.000,ORI_TYP #VAR,CIRC_TYP #BASE,JERK_FAC 50.0000,GEAR_JERK 50.0000,EXAX_IGN 0}
DECL E6POS XP59={X -239.873,Y 70.433,Z 270.000,A -90.001,B 0.123,C 179.669}
DECL FDAT FP59={TOOL_NO 1,BASE_NO 1,IPO_FRAME #BASE,POINT2[] " ",TQ_STATE FALSE}
DECL LDAT LCPDAT59={VEL 0.05000,ACC 100.000,APO_DIST 1.000,APO_FAC 50.0000,AXIS_VEL 100.000,AXIS_ACC 100.000,ORI_TYP #VAR,CIRC_TYP #BASE,JERK_FAC 50.0000,GEAR_JERK 50.0000,EXAX_IGN 0}
DECL E6POS XP60={X -227.408,Y 103.854,Z 270.000,A -90.001,B 0.170,C 179.689}
DECL FDAT FP60={TOOL_NO 1,BASE_NO 1,IPO_FRAME #BASE,POINT2[] " ",TQ_STATE FALSE}
DECL LDAT LCPDAT60={VEL 0.05000,ACC 100.000,APO_DIST 1.000,APO_FAC 50.0000,AXIS_VEL 100.000,AXIS_ACC 100.000,ORI_TYP #VAR,CIRC_TYP #BASE,JERK_FAC 50.0000,GEAR_JERK 50.0000,EXAX_IGN 0}
DECL E6POS XP61={X -210.313,Y 135.160,Z 270.000,A -90.001,B 0.212,C 179.717}
DECL FDAT FP61={TOOL_NO 1,BASE_NO 1,IPO_FRAME #BASE,POINT2[] " ",TQ_STATE FALSE}
DECL LDAT LCPDAT61={VEL 0.05000,ACC 100.000,APO_DIST 1.000,APO_FAC 50.0000,AXIS_VEL 100.000,AXIS_ACC 100.000,ORI_TYP #VAR,CIRC_TYP #BASE,JERK_FAC 50.0000,GEAR_JERK 50.0000,EXAX_IGN 0}
DECL E6POS XP62={X -188.937,Y 163.715,Z 270.000,A -90.001,B 0.250,C 179.750}
DECL FDAT FP62={TOOL_NO 1,BASE_NO 1,IPO_FRAME #BASE,POINT2[] " ",TQ_STATE FALSE}
DECL LDAT LCPDAT62={VEL 0.05000,ACC 100.000,APO_DIST 1.000,APO_FAC 50.0000,AXIS_VEL 100.000,AXIS_ACC 100.000,ORI_TYP #VAR,CIRC_TYP #BASE,JERK_FAC 50.0000,GEAR_JERK 50.0000,EXAX_IGN 0}
DECL E6POS XP63={X -163.715,Y 188.937,Z 270.000,A -90.001,B 0.283,C 179.788}
DECL FDAT FP63={TOOL_NO 1,BASE_NO 1,IPO_FRAME #BASE,POINT2[] " ",TQ_STATE FALSE}
DECL LDAT LCPDAT63={VEL 0.05000,ACC 100.000,APO_DIST 1.000,APO_FAC 50.0000,AXIS_VEL 100.000,AXIS_ACC 100.000,ORI_TYP #VAR,CIRC_TYP #BASE,JERK_FAC 50.0000,GEAR_JERK 50.0000,EXAX_IGN 0}
DECL E6POS XP64={X -135.160,Y 210.313,Z 270.000,A -90.001,B 0.310,C 179.831}
DECL FDAT FP64={TOOL_NO 1,BASE_NO 1,IPO_FRAME #BASE,POINT2[] " ",TQ_STATE FALSE}
DECL LDAT LCPDAT64={VEL 0.05000,ACC 100.000,APO_DIST 1.000,APO_FAC 50.0000,AXIS_VEL 100.000,AXIS_ACC 100.000,ORI_TYP #VAR,CIRC_TYP #BASE,JERK_FAC 50.0000,GEAR_JERK 50.0000,EXAX_IGN 0}
DECL E6POS XP65={X -103.854,Y 227.408,Z 270.000,A -90.001,B 0.332,C 179.876}
DECL FDAT FP65={TOOL_NO 1,BASE_NO 1,IPO_FRAME #BASE,POINT2[] " ",TQ_STATE FALSE}
DECL LDAT LCPDAT65={VEL 0.05000,ACC 100.000,APO_DIST 1.000,APO_FAC 50.0000,AXIS_VEL 100.000,AXIS_ACC 100.000,ORI_TYP #VAR,CIRC_TYP #BASE,JERK_FAC 50.0000,GEAR_JERK 50.0000,EXAX_IGN 0}
DECL E6POS XP66={X -70.433,Y 239.873,Z 270.000,A -90.000,B 0.346,C 179.925}
DECL FDAT FP66={TOOL_NO 1,BASE_NO 1,IPO_FRAME #BASE,POINT2[] " ",TQ_STATE FALSE}
DECL LDAT LCPDAT66={VEL 0.05000,ACC 100.000,APO_DIST 1.000,APO_FAC 50.0000,AXIS_VEL 100.000,AXIS_ACC 100.000,ORI_TYP #VAR,CIRC_TYP #BASE,JERK_FAC 50.0000,GEAR_JERK 50.0000,EXAX_IGN 0}
DECL E6POS XP67={X -35.579,Y 247.455,Z 270.000,A -90.000,B 0.353,C 179.975}
DECL FDAT FP67={TOOL_NO 1,BASE_NO 1,IPO_FRAME #BASE,POINT2[] " ",TQ_STATE FALSE}
DECL LDAT LCPDAT67={VEL 0.05000,ACC 100.000,APO_DIST 1.000,APO_FAC 50.0000,AXIS_VEL 100.000,AXIS_ACC 100.000,ORI_TYP #VAR,CIRC_TYP #BASE,JERK_FAC 50.0000,GEAR_JERK 50.0000,EXAX_IGN 0}
DECL E6POS XP68={X 0.000,Y 250.000,Z 270.000,A -90.000,B 0.353,C 179.975}
DECL FDAT FP68={TOOL_NO 1,BASE_NO 1,IPO_FRAME #BASE,POINT2[] " ",TQ_STATE FALSE}
DECL LDAT LCPDAT68={VEL 0.05000,ACC 100.000,APO_DIST 1.000,APO_FAC 50.0000,AXIS_VEL 100.000,AXIS_ACC 100.000,ORI_TYP #VAR,CIRC_TYP #BASE,JERK_FAC 50.0000,GEAR_JERK 50.0000,EXAX_IGN 0}
DECL E6POS XP69={X 49.895,Y 253.258,Z 319.999,A -90.000,B 0.353,C 179.975}
DECL FDAT FP69={TOOL_NO 1,BASE_NO 1,IPO_FRAME #BASE,POINT2[] " ",TQ_STATE FALSE}
DECL LDAT LCPDAT69={VEL 1.00000,ACC 100.000,APO_DIST 1.000,APO_FAC 50.0000,AXIS_VEL 100.000,AXIS_ACC 100.000,ORI_TYP #VAR,CIRC_TYP #BASE,JERK_FAC 50.0000,GEAR_JERK 50.0000,EXAX_IGN 0}
DECL E6POS XP70={X 49.939,Y 252.642,Z 419.997,A -90.000,B 0.353,C 179.975}
DECL FDAT FP70={TOOL_NO 1,BASE_NO 1,IPO_FRAME #BASE,POINT2[] " ",TQ_STATE FALSE}
DECL LDAT LCPDAT70={VEL 1.00000,ACC 100.000,APO_DIST 1.000,APO_FAC 50.0000,AXIS_VEL 100.000,AXIS_ACC 100.000,ORI_TYP #VAR,CIRC_TYP #BASE,JERK_FAC 50.0000,GEAR_JERK 50.0000,EXAX_IGN 0}
DECL E6AXIS XP71={AXIS: A1 -29.33220,A2 46.67700,A3 -0.02452,A4 26.54560,A5 25.39570,A6 -51.63400}
DECL FDAT FP71={TOOL_NO 1,BASE_NO 1,IPO_FRAME #BASE,POINT2[] " ",TQ_STATE FALSE}
DECL PDAT PPDAT71={VEL 100.000,ACC 100.000,APO_DIST 1.000,GEAR_JERK 50.0000,EXAX_IGN 0}
DECL E6POS XP72={X 187.786,Y 125.499,Z 139.112,A -179.997,B 0.180,C 179.996}
DECL FDAT FP72={TOOL_NO 1,BASE_NO 1,IPO_FRAME #BASE,POINT2[] " ",TQ_STATE FALSE}
DECL LDAT LCPDAT72={VEL 1.00000,ACC 100.000,APO_DIST 1.000,APO_FAC 50.0000,AXIS_VEL 100.000,AXIS_ACC 100.000,ORI_TYP #VAR,CIRC_TYP #BASE,JERK_FAC 50.0000,GEAR_JERK 50.0000,EXAX_IGN 0}
DECL E6POS XP73={X 187.264,Y 125.487,Z 305.356,A 180.000,B 0.184,C -180.000}
DECL FDAT FP73={TOOL_NO 1,BASE_NO 1,IPO_FRAME #BASE,POINT2[] " ",TQ_STATE FALSE}
DECL LDAT LCPDAT73={VEL 1.00000,ACC 100.000,APO_DIST 1.000,APO_FAC 50.0000,AXIS_VEL 100.000,AXIS_ACC 100.000,ORI_TYP #VAR,CIRC_TYP #BASE,JERK_FAC 50.0000,GEAR_JERK 50.0000,EXAX_IGN 0}
DECL E6AXIS XP74={AXIS: A1 -0.00000,A2 0.00000,A3 0.00000,A4 0.00000,A5 0.00000,A6 -0.00000}
DECL FDAT FP74={TOOL_NO 1,BASE_NO 1,IPO_FRAME #BASE,POINT2[] " ",TQ_STATE FALSE}
DECL PDAT PPDAT74={VEL 100.000,ACC 100.000,APO_DIST 1.000,GEAR_JERK 50.0000,EXAX_IGN 0}

ENDDAT
